FUNCTION_BLOCK Distribution2CAT (* CAT Function Block Type *)
  (* Standard: 61499-2 *)
  (* Version 0.0, 7/7/2026, template *)
  PACKAGE Main;
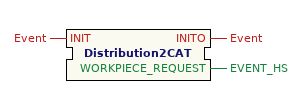
  EVENT_INPUT
    INIT; (* Initialization Request *)
  END_EVENT
  EVENT_OUTPUT
    INITO; (* Initialization Confirm *)
  END_EVENT
  PLUGS
    WORKPIECE_REQUEST : EVENT_HS;
  END_PLUGS
  FBS
    START : E_SR;
    CHECK_STARTED : E_PERMIT;
    FB3 : GiveWorkpiece;
    FB4 : SYMLINKMULTIVARDST_5495E501E675F500(QI := TRUE, NAME1 := '$${PATH}CYL_RET', NAME2 := '$${PATH}CYL_EXT', NAME3 := '$${PATH}WP_PICKED', NAME4 := '$${PATH}ARM_AT_MAG', NAME5 := '$${PATH}ARM_AT_DOWN', NAME6 := '$${PATH}MAG_EMPTY'); {SET_ATTRIBUTE(Configuration.GenericFBType.InterfaceParams, Runtime.System#I:=6;VALUE${I$}:BOOL,BOOL,BOOL,BOOL,BOOL,BOOL)}
    FB5 : SYMLINKMULTIVARSRC_65D63179E2618F5E(QI := TRUE, NAME1 := '$${PATH}VACUUM_ON', NAME2 := '$${PATH}VACCUM_OFF', NAME3 := '$${PATH}ARM_TO_MAG', NAME4 := '$${PATH}ARM_TO_DOWN', NAME5 := '$${PATH}EXTEND_CYL'); {SET_ATTRIBUTE(Configuration.GenericFBType.InterfaceParams, Runtime.System#I:=5;VALUE${I$}:BOOL,BOOL,BOOL,BOOL,BOOL)}
    MagazineCyl : SingleActingCylinder;
    FB7 : ArmReset;
    FB8 : ControlPanel;
    WAIT_WP_INDICATION : E_SR;
    Vacuum : CustomStopActuator;
    Arm : CustomStopActuator;
  END_FBS
  EVENT_CONNECTIONS
    FB4.INITO TO FB5.INIT;
    INIT TO FB4.INIT;
    CHECK_STARTED.EO TO FB3.3D6E8F17A88D01D6;
    WORKPIECE_REQUEST.06D0DEC05BDF54B5 TO CHECK_STARTED.EI;
    FB8.6BF153ECFD1CC9BC TO START.R;
    FB8.C8A63D8D44F6FBE8 TO START.S;
    START.EO TO FB8.94642CF72AED9EF3;
    FB3.4827AB32E389A95A TO Vacuum.B995BB7A7B35D44B;
    FB3.6096B15090B72C95 TO Vacuum.7BAB6103DB1C6BFF;
    FB3.801F2281E3F14364 TO Vacuum.C11C146C3BC053E9;
    FB3.3D7CD2D5BB6105D0 TO WORKPIECE_REQUEST.17D55D3741201415;
    FB3.3D7CD2D5BB6105D0 TO WAIT_WP_INDICATION.R;
    FB3.ED3D348324B91F7E TO WAIT_WP_INDICATION.S;
    FB3.0B9F3017CF4A05C1 TO MagazineCyl.99F4063B254B77CE;
    FB3.A2558C51E8F4B0AC TO MagazineCyl.9F366D7490B55159;
    FB3.D0A914C573069DF6 TO Arm.7BAB6103DB1C6BFF;
    FB3.1B2DEDB9746EFB12 TO Arm.B995BB7A7B35D44B;
    FB3.E0071990EF293838 TO Arm.C11C146C3BC053E9;
    FB5.INITO TO FB8.186CDF42F02DAAF9;
    WAIT_WP_INDICATION.EO TO FB8.D0CE0F6F93E8C4E6;
    FB7.6B9B16A5CCCF0A5F TO FB8.B4AF51BF682610CF;
    FB8.A24AEFFB6D68A233 TO INITO;
    FB8.F94BA7FEBB0FD165 TO FB7.44541FA90B36D44F;
    FB7.4279AF5F2D571F35 TO Arm.B995BB7A7B35D44B;
    FB7.88EB222F28F57D09 TO Arm.7BAB6103DB1C6BFF;
    FB7.AF051DE6AC146B46 TO Arm.C11C146C3BC053E9;
    FB4.CNF TO FB3.7C080AC92CE7241F;
    FB5.INITO TO Vacuum.0250D26CA4B75BF6;
    FB5.INITO TO Arm.0250D26CA4B75BF6;
    FB5.INITO TO MagazineCyl.660CFDEC16C67736;
    Vacuum.30DA918B5EFA21E2 TO FB5.REQ;
    Arm.30DA918B5EFA21E2 TO FB5.REQ;
    MagazineCyl.AB3FD4CE9D9A6580 TO FB5.REQ;
    FB4.CNF TO MagazineCyl.534A07A95E4EF9B6;
    FB4.CNF TO FB7.78E8E2AA9DAF29A8;
  END_CONNECTIONS
  DATA_CONNECTIONS
    FB4.VALUE1 TO FB3.ECF5AB76A8447F7B;
    FB4.VALUE1 TO MagazineCyl.0DA59735E4691A3B;
    FB4.VALUE2 TO MagazineCyl.8562977D9CD64BD4;
    FB4.VALUE2 TO FB3.2C3F87BF27D5CCD5;
    FB4.VALUE4 TO FB3.3CAACAF322D56EE4;
    FB4.VALUE4 TO FB7.4929591747EB6C68;
    FB4.VALUE5 TO FB3.3DE420F02FEBFB11;
    FB4.VALUE5 TO FB7.C845A2BE94918BBD;
    FB4.VALUE6 TO FB3.B13AB1FCC31CCCE4;
    START.Q TO CHECK_STARTED.PERMIT;
    WAIT_WP_INDICATION.Q TO FB8.F66ED9C503CBE986;
    Vacuum.0CAEECB8D3EBC205 TO FB5.VALUE1;
    Vacuum.C60199B3D734C2F9 TO FB5.VALUE2;
    Arm.0CAEECB8D3EBC205 TO FB5.VALUE4;
    Arm.C60199B3D734C2F9 TO FB5.VALUE3;
    MagazineCyl.4D4A774C62CD670B TO FB5.VALUE5;
  END_CONNECTIONS
END_FUNCTION_BLOCK
